(* IEC 61131-3 sources: Test-Git_ESME26/TestProgettoESME_26.fbsproj/PacDriveLib Migration/Motion/Homing/PDL_FB_HomeAbs.fb.st^, 4 files *)

(* ---- AsyncExtDiagTranslation.meth.st ---- *)
METHOD PRIVATE AsyncExtDiagTranslation : BOOL
VAR_INPUT
	i_etResult : SE_Async.ET_Result;
END_VAR

CASE i_etResult OF
	SE_Async.ET_Result.MaxNumOfReusableObjectsExceeded: ; // No error message. Try again to Start in next cycle

	SE_Async.ET_Result.AsyncAddWasNotSuccessful:
		SetDiagOutput(	i_etDiag	:= GD.ET_Diag.UnexpectedProgramBehavior,
						i_etDiagExt := PDL_ET_DiagExt.AsyncAddWasNotSuccessful,
						i_sMsg		:= SE_CTBX.FC_MultiConcat(	i_sString1 := '#',
														i_sString2 := DINT_TO_STRING(diState),
														i_sString3 := ' G_ifAsync.Start: ',
														i_sString4 := PDL_FC_EtDiagExtToString(etDiagExt)));

	SE_Async.ET_Result.InterfaceCastFailed:
		SetDiagOutput(	i_etDiag	:= GD.ET_Diag.UnexpectedProgramBehavior,
						i_etDiagExt := PDL_ET_DiagExt.InterfaceCastFailed,
						i_sMsg		:= SE_CTBX.FC_MultiConcat(	i_sString1 := '#',
														i_sString2 := DINT_TO_STRING(diState),
														i_sString3 := ' G_ifAsync.Start: ',
														i_sString4 := PDL_FC_EtDiagExtToString(etDiagExt)));

	SE_Async.ET_Result.SemaphoreCreateFailed:
		SetDiagOutput(	i_etDiag	:= GD.ET_Diag.UnexpectedProgramBehavior,
						i_etDiagExt := PDL_ET_DiagExt.SemaphoreMeCreateFailed,
						i_sMsg		:= SE_CTBX.FC_MultiConcat(	i_sString1 := '#',
														i_sString2 := DINT_TO_STRING(diState),
														i_sString3 := ' G_ifAsync.Start: ',
														i_sString4 := PDL_FC_EtDiagExtToString(etDiagExt)));

	SE_Async.ET_Result.AsyncInvalid:
		SetDiagOutput(	i_etDiag	:= GD.ET_Diag.InputParameterInvalid,
						i_etDiagExt := PDL_ET_DiagExt.AsyncInvalid,
						i_sMsg		:= SE_CTBX.FC_MultiConcat(	i_sString1 := '#',
														i_sString2 := DINT_TO_STRING(diState),
														i_sString3 := ' G_ifAsync.Start: ',
														i_sString4 := PDL_FC_EtDiagExtToString(etDiagExt)));

	SE_Async.ET_Result.NoAsyncTasksCreated:
		SetDiagOutput(	i_etDiag	:= GD.ET_Diag.ExecutionAborted,
						i_etDiagExt := PDL_ET_DiagExt.NoAsyncTasksCreated,
						i_sMsg		:= SE_CTBX.FC_MultiConcat(	i_sString1 := '#',
														i_sString2 := DINT_TO_STRING(diState),
														i_sString3 := ' G_ifAsync.Start: ',
														i_sString4 := PDL_FC_EtDiagExtToString(etDiagExt)));

	SE_Async.ET_Result.AsyncInitNotFinished:
		SetDiagOutput(	i_etDiag	:= GD.ET_Diag.ExecutionAborted,
						i_etDiagExt := PDL_ET_DiagExt.AsyncInitNotFinished,
						i_sMsg		:= SE_CTBX.FC_MultiConcat(	i_sString1 := '#',
														i_sString2 := DINT_TO_STRING(diState),
														i_sString3 := ' G_ifAsync.Start: ',
														i_sString4 := PDL_FC_EtDiagExtToString(etDiagExt)));

	SE_Async.ET_Result.ColdResetOfControllerNecessary:
		SetDiagOutput(	i_etDiag	:= GD.ET_Diag.ExecutionAborted,
						i_etDiagExt := PDL_ET_DiagExt.ColdResetOfControllerNecessary,
						i_sMsg		:= SE_CTBX.FC_MultiConcat(	i_sString1 := '#',
														i_sString2 := DINT_TO_STRING(diState),
														i_sString3 := ' G_ifAsync.Start: ',
														i_sString4 := PDL_FC_EtDiagExtToString(etDiagExt)));

	ELSE
		SetDiagOutput(	i_etDiag	:= GD.ET_Diag.UnexpectedProgramBehavior,
						i_etDiagExt := PDL_ET_DiagExt.UnexpectedFeedback,
						i_sMsg		:= SE_CTBX.FC_MultiConcat(	i_sString1 := '#',
														i_sString2 := DINT_TO_STRING(diState),
														i_sString3 := ' G_ifAsync.Start: ',
														i_sString4 := PDL_FC_EtDiagExtToString(etDiagExt)));
END_CASE

(* ---- InitInterfaces.meth.st ---- *)
METHOD PRIVATE InitInterfaces : BOOL

VAR
	ifGetParentDevice      : DTSI.IF_GetParentDevice;
	ifDeviceAccess         : DTSI.IF_DeviceAccess;
END_VAR

diSercosState := FC_GetSercosState();

IF diSercosState <> 4 THEN
	SetDiagOutput(	i_etDiag	:= GD.ET_Diag.SercosConditionInvalid,
					i_etDiagExt := PDL_ET_DiagExt.SercosNotInPhaseFour,
					i_sMsg		:= '');
	RETURN;
END_IF

IF i_ifDrive = 0 THEN
	SetDiagOutput(	i_etDiag	:= GD.ET_Diag.InputParameterInvalid,
					i_etDiagExt := PDL_ET_DiagExt.DriveInvalid,
					i_sMsg		:= 'i_ifDrive = 0');
	RETURN;
END_IF

xSuccess := __QUERYINTERFACE(i_ifDrive, ifGetParentDevice);
IF NOT xSuccess OR ifGetParentDevice = 0 THEN
	SetDiagOutput(	i_etDiag	:= GD.ET_Diag.InputParameterInvalid,
					i_etDiagExt := PDL_ET_DiagExt.DriveInvalid,
					i_sMsg		:= 'i_ifDrive - IF_GetParentDevice not implemented.');
	RETURN;
END_IF
ifDeviceAccess := ifGetParentDevice.GetParentDevice();

xSuccess := __QUERYINTERFACE(ifDeviceAccess,ifScalingAccess );
IF (NOT xSuccess OR ifScalingAccess = 0) THEN
	SetDiagOutput(	i_etDiag	:= GD.ET_Diag.InputParameterInvalid,
					i_etDiagExt := PDL_ET_DiagExt.DriveInvalid,
					i_sMsg		:= 'i_ifDrive - IF_Scaling not implemented.');
	RETURN;
END_IF
ifScaling := ifScalingAccess.Scaling;

xSuccess := __QUERYINTERFACE(ifDeviceAccess,ifDrive2Access );
IF (NOT xSuccess OR ifDrive2Access = 0) THEN
	q_etDiag	:= GD.ET_Diag.InputParameterInvalid;
	q_etDiagExt := PDL_ET_DiagExt.DriveInvalid;
	q_sMsg		:= 'i_ifDrive - IF_Drive2 not implemented.';
	RETURN;
END_IF
ifDrive2 := ifDrive2Access.Drive2;

xSuccess := __QUERYINTERFACE(ifDeviceAccess,ifDriveAccess );
IF (NOT xSuccess OR ifDriveAccess = 0) THEN
	q_etDiag	:= GD.ET_Diag.InputParameterInvalid;
	q_etDiagExt := PDL_ET_DiagExt.DriveInvalid;
	q_sMsg		:= 'i_ifDrive - IF_Drive not implemented.';
	RETURN;
END_IF
ifDrive := ifDriveAccess.Drive;

xSuccess := __QUERYINTERFACE(ifDeviceAccess,ifDriveConfigAccess );
IF (NOT xSuccess OR ifDriveConfigAccess = 0) THEN
	SetDiagOutput(	i_etDiag	:= GD.ET_Diag.InputParameterInvalid,
					i_etDiagExt := PDL_ET_DiagExt.DriveInvalid,
					i_sMsg		:= 'i_ifDrive - IF_DriveConfig not implemented.');
	diState := 0;
	RETURN;
END_IF
ifDriveConfig := ifDriveConfigAccess.DriveConfig;

xSuccess := __QUERYINTERFACE(ifDeviceAccess,ifMotorAccess );
IF (NOT xSuccess OR ifMotorAccess = 0) THEN
	SetDiagOutput(	i_etDiag	:= GD.ET_Diag.InputParameterInvalid,
					i_etDiagExt := PDL_ET_DiagExt.DriveInvalid,
					i_sMsg		:= 'i_ifDrive - IF_Motor not implemented.');
	diState := 0;
	RETURN;
END_IF
ifMotor := ifMotorAccess.Motor;

xSuccess := __QUERYINTERFACE(ifDeviceAccess,ifEncoderAccess );
IF (NOT xSuccess OR ifEncoderAccess = 0) THEN
	SetDiagOutput(	i_etDiag	:= GD.ET_Diag.InputParameterInvalid,
					i_etDiagExt := PDL_ET_DiagExt.DriveInvalid,
					i_sMsg		:= 'i_ifDrive - IF_Encoder not implemented.');
	diState := 0;
	RETURN;
END_IF
ifEncoder := ifEncoderAccess.Encoder;

xSuccess := __QUERYINTERFACE(ifDeviceAccess,ifLXM62DriveAccess );
IF (NOT xSuccess OR ifLXM62DriveAccess = 0) THEN
	SetDiagOutput(	i_etDiag	:= GD.ET_Diag.InputParameterInvalid,
					i_etDiagExt := PDL_ET_DiagExt.DriveInvalid,
					i_sMsg		:= 'i_ifDrive - IF_LXM62DriveAccess not implemented.');
	diState := 0;
	RETURN;
END_IF
ifLXM62Drive := ifLXM62DriveAccess.Lexium62Drive;

xSuccess := __QUERYINTERFACE(ifDeviceAccess, ifDeviceType);
IF (NOT xSuccess OR ifDeviceType = 0) THEN
	SetDiagOutput(	i_etDiag	:= GD.ET_Diag.InputParameterInvalid,
					i_etDiagExt := PDL_ET_DiagExt.DriveInvalid,
					i_sMsg 		:= 'i_ifDrive - IF_Device_Type not implemented');
	diState := 0;
	RETURN;
END_IF

InitInterfaces := TRUE;

(* ---- RegisterLoggerPoint.meth.st ---- *)
METHOD PUBLIC RegisterLoggerPoint
VAR_INPUT
	i_ifParent		: APL.IF_LoggerPoint;
	i_sName			: STRING[80];
END_VAR
VAR_OUTPUT
	q_etDiag		: GD.ET_Diag := GD.ET_Diag.Ok;
	q_etDiagExt		: PDL_ET_DiagExt := PDL_ET_DiagExt.Ok;
END_VAR
VAR
	etDiagBuffer		: GD.ET_Diag;
	etDiagExtBufferAPL	: APL.ET_DiagExt;
END_VAR

THIS^.fbLoggerPoint.RegisterLoggerPoint(	i_ifParent		:= i_ifParent,
											i_sName			:= i_sName,
											i_sType			:= 'FB_HomeAbs',
											i_sSource		:= 'PDL',
											q_etDiag		=> etDiagBuffer,
											q_etDiagExt		=> etDiagExtBufferAPL);
IF (etDiagBuffer <> GD.ET_Diag.Ok) THEN
	CASE etDiagExtBufferAPL OF
		APL.ET_DiagExt.ParentInvalid:
			q_etDiag := GD.ET_Diag.InputParameterInvalid;
			q_etDiagExt := PDL_ET_DiagExt.ParentInvalid;

		APL.ET_DiagExt.ParentNotRegistered:
			q_etDiag := GD.ET_Diag.InputParameterInvalid;
			q_etDiagExt := PDL_ET_DiagExt.ParentNotRegistered;

		APL.ET_DiagExt.MaxNumberOfLoggerPointsExeeded:
			q_etDiag := GD.ET_Diag.InputParameterInvalid;
			q_etDiagExt := PDL_ET_DiagExt.MaxNumberOfLoggerPointsExeeded;

	ELSE
		q_etDiag := GD.ET_Diag.UnexpectedProgramBehavior;
		q_etdiagExt := PDL_ET_DiagExt.UnexpectedDiagExt;
	END_CASE
END_IF

(* ---- SetDiagOutput.meth.st ---- *)
METHOD PRIVATE SetDiagOutput : BOOL
VAR_INPUT
	i_etDiag	: GD.ET_Diag;
	i_etDiagExt	: PDL_ET_DiagExt;
	i_sMsg		: STRING[80];
END_VAR
VAR
END_VAR

IF i_etDiag <> GD.ET_Diag.Ok THEN
	q_xBusy := FALSE;
	q_xReady := FALSE;
END_IF
IF q_etDiag = GD.ET_Diag.OK OR i_etDiagExt = PDL_ET_DiagExt.Disabled THEN
	q_etDiag := i_etDiag;
	q_etDiagExt := i_etDiagExt;
	q_sMsg := i_sMsg;

	IF(i_etDiag = GD.ET_Diag.Ok) AND (THIS^.fbLoggerPoint.etLogLevel >= APL.ET_LogLevel.StatusMessage) THEN
		THIS^.fbLoggerPoint.AddLogEntry(	i_etLogLevel	:= APL.ET_LogLevel.StatusMessage,
											i_etDiag		:= q_etDiag,
											i_udiDiagExt	:= q_etDiagExt,
											i_sMessage		:= SE_CTBX.FC_MultiConcat(	i_sString1	:= Standard.CONCAT('ET_Diag: ', GD.FC_EtDiagToString(q_etDiag)),
																				i_sString2	:= Standard.CONCAT(' PDL_ET_DiagExt: ', PDL_FC_EtDiagExtToString(q_etDiagExt)),
																				i_sString3	:= Standard.CONCAT(' sMsg: ', q_sMsg),
																				i_sString4	:= ''),
											q_etDiag		:= ,	// ignore result
											q_etDiagExt		:= );	// ignore result
	ELSIF(i_etDiag = GD.ET_Diag.UnexpectedProgramBehavior) AND (THIS^.fbLoggerPoint.etLogLevel >= APL.ET_LogLevel.CriticalException) THEN
		THIS^.fbLoggerPoint.AddLogEntry(	i_etLogLevel	:= APL.ET_LogLevel.CriticalException,
											i_etDiag		:= q_etDiag,
											i_udiDiagExt	:= q_etDiagExt,
											i_sMessage		:= SE_CTBX.FC_MultiConcat(	i_sString1	:= Standard.CONCAT('ET_Diag: ', GD.FC_EtDiagToString(q_etDiag)),
																				i_sString2	:= Standard.CONCAT(' PDL_ET_DiagExt: ', PDL_FC_EtDiagExtToString(q_etDiagExt)),
																				i_sString3	:= Standard.CONCAT(' sMsg: ', q_sMsg),
																				i_sString4	:= ''),
											q_etDiag		:= ,	// ignore result
											q_etDiagExt		:= );	// ignore result
	ELSIF(i_etDiag <> GD.ET_Diag.Ok) AND (THIS^.fbLoggerPoint.etLogLevel >= APL.ET_LogLevel.Exception) THEN
		THIS^.fbLoggerPoint.AddLogEntry(	i_etLogLevel	:= APL.ET_LogLevel.Exception,
											i_etDiag		:= q_etDiag,
											i_udiDiagExt	:= q_etDiagExt,
											i_sMessage		:= SE_CTBX.FC_MultiConcat(	i_sString1	:= Standard.CONCAT('ET_Diag: ', GD.FC_EtDiagToString(q_etDiag)),
																				i_sString2	:= Standard.CONCAT(' PDL_ET_DiagExt: ', PDL_FC_EtDiagExtToString(q_etDiagExt)),
																				i_sString3	:= Standard.CONCAT(' sMsg: ', q_sMsg),
																				i_sString4	:= ''),
											q_etDiag		:= ,	// ignore result
											q_etDiagExt		:= );	// ignore result
	END_IF
END_IF
